(* IEC 61131-3 sources: Versio-VersionControlSystem/fixtures/projects/TC3_PlcSample_reStrText/TC3_PlcSample_reStrText/LibraryDocumentationSample Project/LibPOUs/B_DocuElements/Lists, 4 files *)

(* ---- FB_Libdoc_DefinitionList.st ---- *)
(*
Term 1
    Definition 1.

Term 2
    Definition 2, paragraph 1.

    Definition 2, paragraph 2.

Term 3 : classifier
    Definition 3.

Term 4 : classifier one : classifier two
    - Item 1
    - Item 2
*)

FUNCTION_BLOCK FB_Libdoc_DefinitionList
VAR_INPUT
    nVarA : INT;
    nVarB : INT;
END_VAR
VAR_OUTPUT
    nSum : INT;
END_VAR
VAR
END_VAR

(* ---- FB_Libdoc_FieldList.st ---- *)
(*
:Organization: Beckhoff Automation GmbH & Co. KG
:Contact: info@beckhoff.de
:Address: | Hülshorstweg 20
          | 33415 Verl
          | Germany
:Authors: - Me
          - Myself
          - I
:Version: 1.0
:Status: released
:Date: 2017-12-07

:Copyright:
 © Beckhoff Automation GmbH & Co. KG, Germany.
 The reproduction, distribution and utilization of this document as well as
 the communication of its contents to others without express authorization are prohibited.
 Offenders will be held liable for the payment of damages.
 All rights reserved in the event of the grant of a patent, utility model or design.
:Abstract: topic
:Indentation:
 Since the field marker may be quite long, the second
 and subsequent lines of the field body do not have to line up
 with the first line, but they must be indented relative to the
 field name marker, and they must line up with each other.
:LongLongFieldname: Since the field marker is quite long,
                    the field body is shown in the line after the marker.
:Parameter nIn: Integer
:Parameter nVarB: Integer
:*Parameter nVarC*: Integer
:``Parameter nVarD``: Integer
*)

FUNCTION_BLOCK FB_Libdoc_FieldList
VAR_INPUT
    nVarA : INT;
    nVarB : INT;
END_VAR
VAR_OUTPUT
    nSum : INT;
END_VAR
VAR
END_VAR

(* ---- FB_Libdoc_OrderedNumberedEnumerationList.st ---- *)
(*
1) This is the first item in the list.

   (a) This is the first subitem (1a).
   (b) This is the second subitem (1b).

2) This is the second item in the list.

   (a) This is the first subitem (2a).
   (b) This is the second subitem (2b).

#) This item is auto-enumerated.
*)

FUNCTION_BLOCK FB_Libdoc_OrderedNumberedEnumerationList
VAR_INPUT
    nVarA : INT;
    nVarB : INT;
END_VAR
VAR_OUTPUT
    nSum : INT;
END_VAR
VAR
END_VAR

(* ---- FB_Libdoc_UnorderedEnumerationList.st ---- *)
(*
This paragraph is not part of the list.

- This is the first bullet list item.  The blank line above the
  first list item is required; blank lines between list items
  (such as below this paragraph) are optional.

  - This is a sublist. The bullet lines up with the left edge
    of the text blocks above. A sublist is a new list so
    requires a blank line above. A blank line below is optional.

  - This is a sublist. The bullet lines up with the left edge
    of the text blocks above. A sublist is a new list so
    requires a blank line above. A blank line below is optional.

- This is the second item of the main list.

- This is the third item of the main list.

This paragraph is not part of the list.
*)

FUNCTION_BLOCK FB_Libdoc_UnorderedEnumerationList
VAR_INPUT
    nVarA : INT;
    nVarB : INT;
END_VAR
VAR_OUTPUT
    nSum : INT;
END_VAR
VAR
END_VAR
